// TwinCAT 3 PLC project Lab_02
// ProgramVersion: 3.1.4026.27
// libraries:
//   Tc2_Standard, * (Beckhoff Automation GmbH)
//   Tc2_System, * (Beckhoff Automation GmbH)
// project tree:
//   GVLs/ IN_OUT.TcGVL
//   / PlcTask.TcTTO
//   POUs/ MAIN.TcPOU
// real-time tasks:
//   TASK PlcTask: cycle T#10ms, priority 20, ADS port 350
// I/O:
//   DEVICE Gerät 1 (EtherCAT), AmsNetId 199.4.42.250.2.1
//     Box 1 (EPP2316-0003) [EPP2316-0003 8 K. Dig. Ein, 10µs, 8 K. Dig. Aus 24V, 0,5A, Diagnose, 10-Pol Steckverbinder]
// variable links:
//   Lab_02/Lab_02 Instance <-> Device 1 (EtherCAT)/Box 1 (EPP2316-0003)
//     PlcTask Inputs/IN_OUT._i_b_endSwitch_{1..4} <-> DIG Inputs/Input {1..4}  (4 links)
//     PlcTask Inputs/IN_OUT._i_b_startButton <-> DIG Inputs/Input 5
//     PlcTask Inputs/IN_OUT._i_b_stopButton <-> DIG Inputs/Input 6
//     PlcTask Outputs/IN_OUT._o_b_valve{1..4} <-> DIG Outputs/Output {1..4}  (4 links)

CONFIGURATION Lab_02
    RESOURCE PLC ON TwinCAT3
        TASK PlcTask(INTERVAL := T#10ms, PRIORITY := 20);
        PROGRAM MAIN WITH PlcTask : MAIN;
    END_RESOURCE
END_CONFIGURATION

// ---- GVLs/IN_OUT.TcGVL
{attribute 'qualified_only'}
VAR_GLOBAL
	
	_i_b_endSwitch_1 AT %I* :BOOL;
	_i_b_endSwitch_2 AT %I* :BOOL;
	_i_b_endSwitch_3 AT %I* :BOOL;
	_i_b_endSwitch_4 AT %I* :BOOL;
	_i_b_startButton AT %I*	:BOOL;
	_i_b_stopButton	 AT %I*	:BOOL;

	_o_b_valve1	AT %Q*	:BOOL;
	_o_b_valve2	AT %Q*	:BOOL;
	_o_b_valve3	AT %Q*	:BOOL;
	_o_b_valve4	AT %Q*	:BOOL;



END_VAR

// ---- POUs/MAIN.TcPOU
PROGRAM MAIN
VAR
	l_b_step :INT;
	l_flankeStartbutton : R_TRIG;
	
	l_i_counter :INT;
END_VAR

l_flankeStartbutton(CLK := IN_OUT._i_b_startButton);

IF NOT IN_OUT._i_b_stopButton OR l_i_counter = 3 THEN
	l_b_step := 100;
END_IF

CASE l_b_step OF
	0:
		IF l_flankeStartbutton.Q AND IN_OUT._i_b_endSwitch_3 AND IN_OUT._i_b_endSwitch_1 AND IN_OUT._i_b_stopButton THEN
			l_b_step := 1;
		END_IF
	1:
		IN_OUT._o_b_valve1 := TRUE;
		IF IN_OUT._i_b_endSwitch_2 THEN
			IN_OUT._o_b_valve1 := FALSE;
			l_b_step := 2;
		END_IF
	2: 
		IN_OUT._o_b_valve2 := TRUE;
		IF IN_OUT._i_b_endSwitch_1 THEN
			IN_OUT._o_b_valve2 := FALSE;
			l_b_step := 3;
		END_IF
	3:
		IN_OUT._o_b_valve3 := TRUE;
		IF IN_OUT._i_b_endSwitch_4 THEN
			IN_OUT._o_b_valve3 := FALSE;
			l_b_step := 4;
		END_IF
	4: 
		IN_OUT._o_b_valve4 := TRUE;
		IF IN_OUT._i_b_endSwitch_3 THEN
			l_i_counter := l_i_counter +1;
			IN_OUT._o_b_valve4 := FALSE;
			l_b_step := 1;
		END_IF
	100:
		IN_OUT._o_b_valve1 := TRUE;
		IN_OUT._o_b_valve3 := TRUE;
		l_i_counter := 0;
		
		IF IN_OUT._i_b_endSwitch_1 THEN
			IN_OUT._o_b_valve1 := FALSE;
		END_IF
		
		IF IN_OUT._i_b_endSwitch_3 THEN
			IN_OUT._o_b_valve3 := FALSE;
		END_IF
		
		IF IN_OUT._i_b_endSwitch_1 AND IN_OUT._i_b_endSwitch_3 THEN
			l_b_step := 0;
		END_IF
END_CASE

END_PROGRAM
